Staubli VAL3: LibTorque.pjx

--- LibTorque.pjx ---
Parameters version=s8.15.3Cs9_BS3337 stackSize=5000 millimeterUnit=true
Program file=_getSetForce.pgx
Program file=_setMaxJntForce.pgx
Program file=getArmTypeList.pgx
Program file=initParameter.pgx
Program file=readme.pgx
Program file=refresh.pgx
Program file=setPageMaxJntForce.pgx
Program file=start.pgx
Program file=stop.pgx
Program file=unLock.pgx
Data file=LibTorque.dtx
Library alias=forcedata path=./data/ForceData/ForceData.pjx

--- LibTorque.dtx ---
public bool bDisable[4]
  [0] = true
  [1] = true
  [2] = true
  [3] = true
bool bLock
bool bSix_Axis
mdesc mNomSpeed
num nCurrentMaxForce
public num nMaxJntForce[4]
  [0] = 1000000
  [1] = 1000000
  [2] = 21.1
  [3] = 65
num nMaxJntGet
string sArm4List[9]
  [0] = "tp_80"
  [1] = "ts2_100"
  [2] = "ts2_40"
  [3] = "ts2_60"
  [4] = "ts2_80"
  [5] = "ts_20"
  [6] = "ts_40"
  [7] = "ts_60"
  [8] = "ts_80"
string sArm6List[16]
  [0] = "rx_160"
  [1] = "tx2_140"
  [2] = "tx2_160"
  [3] = "tx2_160l"
  [4] = "tx2_200"
  [5] = "tx2_200l"
  [6] = "tx2_40"
  [7] = "tx2_60"
  [8] = "tx2_60l"
  [9] = "tx2_90"
  [10] = "tx2_90l"
  [11] = "tx2_90xl"
  [12] = "tx_200"
  [13] = "tx_40"
  [14] = "tx_60"
  [15] = "tx_90"
string sArmDetail = "ts2_40"
string sArmType = "4_Axis"
public string sBtnUnLock = "保存"
string sPassword = "staubli2025"

--- start.pgx ---
program start()
begin
end

--- _getSetForce.pgx ---
public program _getSetForce(num& x_nCurrentMaxForce[], string& x_sKey, string& x_sArmType, bool& x_bFind)
// 功能：获取对应型号机器人设定的扭矩限值
// //x_nCurrentMaxForce 当前机型扭矩库设置的最大限值
// //x_sKey   扭矩库键值
// //x_sArmType 反馈四轴/六轴机器人
// //x_bFind 是否在扭矩库中找到当前机型
  local string l_sArmType
  local num i
  local bool l_bIsScara
begin
  //x_nCurrentMaxForce 当前机型扭矩库设置的最大限值
  //x_sKey             扭矩库键值
  //x_sArmType         反馈四轴/六轴机器人
  //x_bFind            是否在扭矩库中找到当前机型
  x_bFind=false
  //获取对应型号机器人设定的扭矩限值
  //获取机器人型号
  l_sArmType=getVersion("Arm Type")
  //打印机器人型号
  logMsg(l_sArmType)
  l_bIsScara=(left(l_sArmType,2)=="rs" or left(l_sArmType,2)=="ts" or left(l_sArmType,2)=="tp")
  l_sArmType=left(l_sArmType,find(l_sArmType,"-"))
  call getArmTypeList(sArm4List,sArm6List)
  //判断机器人4轴/6轴
  if l_bIsScara
    //获取机器人扭矩设定值
    for i=0 to size(sArm4List)-1
      if l_sArmType==sArm4List[i]
        resize(x_nCurrentMaxForce,1,4)
        x_nCurrentMaxForce[0]=forcedata:tArm4Force[sArm4List[i]].nMaxJnt4Force[0]
        x_nCurrentMaxForce[1]=forcedata:tArm4Force[sArm4List[i]].nMaxJnt4Force[1]
        x_nCurrentMaxForce[2]=forcedata:tArm4Force[sArm4List[i]].nMaxJnt4Force[2]
        x_nCurrentMaxForce[3]=forcedata:tArm4Force[sArm4List[i]].nMaxJnt4Force[3]
        x_sKey=l_sArmType
        x_sArmType="4_Axis"
        x_bFind=true
      endIf
    endFor
  else
    for i=0 to size(sArm6List)-1
      if l_sArmType==sArm6List[i]
        resize(x_nCurrentMaxForce,1,6)
        x_nCurrentMaxForce[0]=forcedata:tArm6Force[sArm6List[i]].nMaxJnt6Force[0]
        x_nCurrentMaxForce[1]=forcedata:tArm6Force[sArm6List[i]].nMaxJnt6Force[1]
        x_nCurrentMaxForce[2]=forcedata:tArm6Force[sArm6List[i]].nMaxJnt6Force[2]
        x_nCurrentMaxForce[3]=forcedata:tArm6Force[sArm6List[i]].nMaxJnt6Force[3]
        x_nCurrentMaxForce[4]=forcedata:tArm6Force[sArm6List[i]].nMaxJnt6Force[4]
        x_nCurrentMaxForce[5]=forcedata:tArm6Force[sArm6List[i]].nMaxJnt6Force[5]
        x_sKey=l_sArmType
        x_sArmType="6_Axis"
        x_bFind=true
      endIf
    endFor
  endIf

end

--- _setMaxJntForce.pgx ---
public program _setMaxJntForce()
// //设置机器人各个轴扭矩最大值
  local bool l_bFind
  local num i
  local string l_sKey
begin
  //根据型号获取扭矩限制值
  call _getSetForce(nCurrentMaxForce,sArmDetail,sArmType,l_bFind)
  if l_bFind
    for i=0 to size(nCurrentMaxForce)-1
      logMsg(l_sKey+" J"+toString("",i+1)+"设定限制："+toString("",nCurrentMaxForce[i]))
    endFor
    //设置机器人各个轴最大扭矩
    $setMaxJntForce(nCurrentMaxForce)
    delay(0.5)
    //手臂实际扭矩限制值
    resize(nMaxJntGet,1,size(nCurrentMaxForce))
    $getMaxJntForce(nMaxJntGet)
    for i=0 to size(nMaxJntGet)-1
      logMsg(l_sKey+" J"+toString("",i+1)+"实际限制："+toString("",nMaxJntGet[i]))
    endFor
  else
    logMsg("扭矩库中缺少当前机器人型号，请添加!!!")
  endIf
end

--- getArmTypeList.pgx ---
public program getArmTypeList(string& x_sItem[], string& x_sItem2[])
// //获取所有4轴6轴机器人型号列表
// //x_sItem  4轴手臂型号列表
// //x_sItem2 6轴手臂型号列表
  local trsf l_tTrsf
  local string l_sItem[6]
  local string l_sEvent
  local string l_sItem2[7]
  local string l_sKey[2]
  local num i
  local num j
begin
  //获取所有4轴6轴机器人型号列表
  //x_sItem  4轴手臂型号列表
  //x_sItem2 6轴手臂型号列表
  //获取列表
  resize(x_sItem,1,size(forcedata:tArm4Force))
  resize(x_sItem2,1,size(forcedata:tArm6Force))
  l_sKey=first(forcedata:tArm4Force)
  l_sKey[1]=first(forcedata:tArm6Force)
  i=0
  j=0
  while l_sKey!=""
    x_sItem[i]=l_sKey
    l_sKey=next(forcedata:tArm4Force[l_sKey])
    i=i+1
  endWhile
  while l_sKey[1]!=""
    x_sItem2[j]=l_sKey[1]
    l_sKey[1]=next(forcedata:tArm6Force[l_sKey[1]])
    j=j+1
  endWhile
  if l_sKey=="" and i==0
    x_sItem[i]=""
  endIf
  if l_sKey[1]=="" and j==0
    x_sItem2[j]=""
  endIf
end

--- initParameter.pgx ---
public program initParameter()
  local string l_sKey
  local bool l_bFind
  local num i
begin
  //功能：设置扭矩限值界面初始化调用
  bLock=true
  sBtnUnLock="解锁"
  //获取机器人类型
  call _getSetForce(nMaxJntForce,sArmDetail,sArmType,l_bFind)
  if l_bFind
    if sArmType=="4_Axis"
      resize(bDisable,1,4)
      //resize(nMaxJntForce,1,4)
      bSix_Axis=false
    elseIf sArmType=="6_Axis"
      resize(bDisable,1,6)
      //resize(nMaxJntForce,1,6)
      userPageBind("setJntForce","nmb1_Copy3","disabled",bDisable[4],1,"r")
      userPageBind("setJntForce","nmb1_Copy3","value",nMaxJntForce[4],1,"rw")
      userPageBind("setJntForce","nmb1_Copy5","disabled",bDisable[5],1,"r")
      userPageBind("setJntForce","nmb1_Copy5","value",nMaxJntForce[5],1,"rw")
      bSix_Axis=true
    endIf
    //初始化扭矩设置解锁按钮
    for i=0 to size(bDisable)-1
      bDisable[i]=true
    endFor
  else
    logMsg("扭矩库中缺少当前机器人型号，请添加!!!")
  endIf
end

--- readme.pgx ---
program readme()
begin
  //2025.04.15
  //该库用于获取机器人对应机型设置的各个关节轴的最大扭矩值
  //_getSetForce 功能：获取扭矩库存放机型各个轴关节扭矩限值
  //_setMaxJntForce 功能：设置对应机型各个轴关节扭矩限值
  //getArmTypeList 功能：获取扭矩库机型名称列表
  //initParameter 功能：设置扭矩限值界面初始化调用
  //setPageMaxJntForce 功能：页面修改扭矩库限值
  //refresh 功能：设置扭矩限值界面实时刷新调用
  //unLock 功能：设置扭矩限值界面解锁按钮调用

  //---------------------------示例---------------------------------//
  //   //初始化调用
  //  call libtqe:initParameter()
  //   //设置扭矩限值界面（自定义）
  //  userPage("new1")
  //  do

  //    //刷新解锁/保存按钮
  //    call libtqe:refresh()
  //    delay(0)
  //  until false
end

--- refresh.pgx ---
public program refresh()
begin
  //功能：设置扭矩限值界面实时刷新调用
  if bLock==true
    sBtnUnLock="解锁"
  else
    sBtnUnLock="保存"
  endIf
end

--- setPageMaxJntForce.pgx ---
public program setPageMaxJntForce()
  local num i
begin
  //页面修改扭矩库限值
  if sArmType=="4_Axis"
    for i=0 to 3
      forcedata:tArm4Force[sArmDetail].nMaxJnt4Force[i]=nMaxJntForce[i]
    endFor
  elseIf sArmType=="6_Axis"
    for i=0 to 5
      forcedata:tArm6Force[sArmDetail].nMaxJnt6Force[i]=nMaxJntForce[i]
    endFor
  endIf
  forcedata:libSave()
  delay(0.1)
end

--- stop.pgx ---
program stop()
begin
end

--- unLock.pgx ---
public program unLock()
  local string l_sEntry
  local bool l_bResult
  local num i
  local bool l_bFind
begin
  if bLock==true
    l_bResult=userPagePrompt("请输入密码",l_sEntry)
    if l_bResult==false
      return
    endIf
    if l_sEntry!=sPassword[0]
      popUpMsg("密码错误")
      return
    endIf
    //2024.04.29 add解锁扭矩限位设置
    for i=0 to size(bDisable)-1
      bDisable[i]=false
    endFor
    popUpMsg("修改后请点击保存!")
    bLock=false
  else
    for i=0 to size(bDisable)-1
      bDisable[i]=true
    endFor
    call setPageMaxJntForce()
    call _getSetForce(nMaxJntForce,sArmDetail,sArmType,l_bFind)
    popUpMsg("机器人关节扭矩限制保存成功!")
    bLock=true
  endIf
end
